Fanuc KAREL source: KT00718.KL

PROGRAM KT00718
%NOLOCKGROUP
VAR
  P1: POSITION
  P2: POSITION
  OUT: BOOLEAN
BEGIN
  OUT = UNINIT(P1)
END KT00718
